Fanuc KAREL source: kf00080.KL

-- PROVISIONAL review KL for V940-1; original PC SHA256 af125d89c5f51b11d897a9c294691aa594924dbc1b0a872fcf26c90daf27956c
-- Incomplete behavior may be omitted. Consult companion uncertainty JSON. Do not deploy.
PROGRAM KF00080
%NOLOCKGROUP
BEGIN
  -- V9_ZERO_TABLE_METADATA_HINT layout=0002_ascii; no indexed target words; source/name/runtime held
  -- UNRESOLVED_PC offsets 5-15; opcodes 27,22,31
  -- UNRESOLVED_PC offsets 20-24; opcodes 7F
END KF00080
